FUNCTION_BLOCK OBSTACLE_AVOID (* E-puck obstacle avoidance fb *)
  (* Standard: 61499-2; Classification: Basic; ApplicationDomain: Robotics; Function: Navigation; Type: Basic; Description: E-puck obstacle avoidance FB *)
  (* Version 1.0, 2026-10-22, Mauricio Martins Taques Filho, GASR/UDESC, Initial version *)
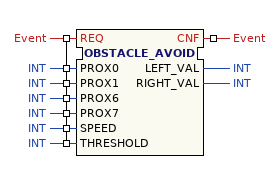
  EVENT_INPUT
    REQ WITH PROX0, PROX1, PROX6, PROX7, SPEED, THRESHOLD; (* Pace determiner *)
  END_EVENT
  EVENT_OUTPUT
    CNF WITH LEFT, RIGHT; (* Determined pace *)
  END_EVENT
  VAR_INPUT
    PROX0 : INT; (* Upper right sensor *)
    PROX1 : INT; (* Right/front sensor *)
    PROX6 : INT; (* Left/front sensor *)
    PROX7 : INT; (* Upper left sensor *)
    SPEED : INT := 500; (* Robot speed in steps *)
    THRESHOLD : INT := 1000; (* Limit sensor value *)
  END_VAR
  VAR_OUTPUT
    LEFT_VAL : INT; (* Left wheel pace *)
    RIGHT_VAL : INT; (* Right wheel pace *)
  END_VAR
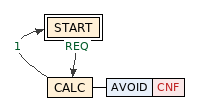
  EC_STATES
    START; (* Initial State *)
    CALC : AVOID -> CNF;
  END_STATES
  EC_TRANSITIONS
    START TO CALC := REQ;
    CALC TO START := 1;
  END_TRANSITIONS
  ALGORITHM AVOID IN ST: (* Moves to the side opposite the obstacle *)
IF PROX0 + PROX1 > THRESHOLD THEN
    LEFT_VAL := -SPEED / 2;
    RIGHT_VAL := SPEED / 2;
ELSIF PROX6 + PROX7 > THRESHOLD THEN
    LEFT_VAL := SPEED / 2;
    RIGHT_VAL := -SPEED / 2;
ELSE
    LEFT_VAL := SPEED;
    RIGHT_VAL := SPEED;
END_IF;
  END_ALGORITHM
END_FUNCTION_BLOCK
